Fanuc KAREL source: KB00070.KL

PROGRAM KB00070
%NOLOCKGROUP
%ENVIRONMENT ERRS
VAR
  P1: INTEGER
  P2: INTEGER
  P3: STRING[80]
  P4: INTEGER
  P5: STRING[80]
  P6: INTEGER
  P7: INTEGER
  P8: STRING[80]
BEGIN
  P1 = 1
  P2 = 1
  P3 = 'A'
  P4 = 1
  P5 = 'A'
  P6 = 1
  P7 = 1
  P8 = 'A'
  ERR_DATA(P1, P2, P3, P4, P5, P6, P7, P8)
END KB00070
